Fanuc KAREL source: KT00985.KL

PROGRAM KT00985
%NOLOCKGROUP
VAR
  Y1: ARRAY[2] OF BYTE
  Y2: ARRAY[2] OF BYTE
  CFG: CONFIG
  OUT: POSITION
BEGIN
  Y1[1] = 2
  Y2[1] = 3
  Y1[1] = 2
  Y2[1] = 3
  CFG.CFG_FLIP = TRUE
  OUT = POS(Y1[1], Y1[1], Y1[1], Y1[1], Y1[1], Y1[1], CFG)
END KT00985
